(* IEC 61131-3 sources: FACTORY_io/fabrica-viva/etapa-6, 3 files *)

(* ---- fragmento-bloques.st ---- *)
(* ===== Etapa 6 · Bloque de función FB_Muting =====
   La cortina del muelle protege a las personas: si algo la corta, la línea se para. Pero los palés
   tienen que pasar por ella. El muting la anula solo mientras pasa un palé:
   - Empieza si los dos sensores de muting se tapan en orden: primero A y después B (el flanco de
     subida de B con A tapado). Una persona que cruza la cortina no los tapa así.
   - Acaba cuando la carga ha pasado: A y B libres y la cortina despejada.
   - Por seguridad, como mucho 30 s seguidos.
   ZonaSegura := la cortina libre, o el muting activo. *)
FUNCTION_BLOCK FB_Muting
VAR_INPUT
  SensorA : BOOL;       (* sensor de muting antes de la cortina *)
  SensorB : BOOL;       (* sensor de muting, más cerca de la cortina *)
  CortinaLibre : BOOL;  (* salida de seguridad de la cortina: TRUE = nada la corta *)
END_VAR
VAR_OUTPUT
  Activo : BOOL;        (* el muting está anulando la cortina *)
  ZonaSegura : BOOL;    (* se puede trabajar *)
END_VAR
VAR
  (* tus variables internas del bloque *)
END_VAR

(* ---- tu código del bloque ---- *)
END_FUNCTION_BLOCK

(* ---- solucion.st ---- *)
(* Fábrica viva · Etapa 6 · Solución de referencia: enfardado, expedición y cortina de seguridad con muting. *)
FUNCTION_BLOCK FB_Cola
VAR_INPUT
  Meter : BOOL;
  Valor : DINT;
  Sacar : BOOL;
END_VAR
VAR_OUTPUT
  Primero : DINT;
  Cantidad : INT;
END_VAR
VAR
  Datos : ARRAY[0..15] OF DINT;
  i : INT;
END_VAR

(* Sacar desplaza todo un puesto hacia la cabeza; meter escribe detrás del último. *)
IF Sacar AND Cantidad > 0 THEN
  FOR i := 0 TO 14 DO
    Datos[i] := Datos[i + 1];
  END_FOR;
  Cantidad := Cantidad - 1;
END_IF;
IF Meter AND Cantidad < 16 THEN
  Datos[Cantidad] := Valor;
  Cantidad := Cantidad + 1;
END_IF;
IF Cantidad > 0 THEN
  Primero := Datos[0];
ELSE
  Primero := 0;
END_IF;
END_FUNCTION_BLOCK

FUNCTION_BLOCK FB_Muting
VAR_INPUT
  SensorA : BOOL;
  SensorB : BOOL;
  CortinaLibre : BOOL;
END_VAR
VAR_OUTPUT
  Activo : BOOL;
  ZonaSegura : BOOL;
END_VAR
VAR
  SubeB : R_TRIG;
  Limite : TON;
END_VAR

(* El muting empieza solo si los dos sensores se tapan en orden, A y luego B, como hace un palé al
   llegar; una persona que cruza la cortina no los tapa así. Acaba cuando la carga ha pasado: los dos
   sensores libres y la cortina despejada. Con un tiempo máximo, por si se queda algo a medias. *)
SubeB(CLK := SensorB);
IF SubeB.Q AND SensorA THEN
  Activo := TRUE;
END_IF;
IF Activo AND NOT SensorA AND NOT SensorB AND CortinaLibre THEN
  Activo := FALSE;
END_IF;
Limite(IN := Activo, PT := T#30s);
IF Limite.Q THEN
  Activo := FALSE;
END_IF;
ZonaSegura := CortinaLibre OR Activo;
END_FUNCTION_BLOCK

FUNCTION_BLOCK FB_Paletizado
VAR_INPUT
  Habilitar : BOOL;
  CajaLista : BOOL;
  PaleListo : BOOL;
  RobotListo : BOOL;
  Reiniciar : BOOL;
END_VAR
VAR_OUTPUT
  Trabajo : INT;
  Ejecutar : BOOL;
  Paso : INT;
  Colocadas : INT;
  Total : INT;
  PaleLleno : BOOL;
END_VAR

(* Intercambio de señales con el robot: se fija el trabajo, se mantiene Ejecutar hasta que el robot
   avisa de que lo ha empezado (cae RobotListo) y se espera a que vuelva a estar listo. *)
Ejecutar := FALSE;
CASE Paso OF
  0: (* esperando caja y palé *)
    IF Reiniciar THEN
      Colocadas := 0;
    END_IF;
    IF Habilitar AND CajaLista AND PaleListo AND RobotListo AND Colocadas < 8 THEN
      Trabajo := 1;
      Paso := 1;
    END_IF;
  1: (* recoger: orden dada *)
    Ejecutar := TRUE;
    IF NOT RobotListo THEN
      Paso := 2;
    END_IF;
  2: (* recogiendo *)
    IF RobotListo AND Habilitar THEN
      Trabajo := 2 + Colocadas;
      Paso := 3;
    END_IF;
  3: (* dejar en su hueco: orden dada *)
    Ejecutar := TRUE;
    IF NOT RobotListo THEN
      Paso := 4;
    END_IF;
  4: (* dejando y volviendo a reposo *)
    IF RobotListo THEN
      Colocadas := Colocadas + 1;
      Total := Total + 1;
      Paso := 0;
    END_IF;
END_CASE;
PaleLleno := Colocadas >= 8;
END_FUNCTION_BLOCK

FUNCTION_BLOCK FB_Pulmon
VAR_INPUT
  Habilitar : BOOL;
  CajaEnTope : BOOL;
  Permiso : BOOL;
END_VAR
VAR_OUTPUT
  Tope : BOOL;
  Avance : BOOL;
  Salida : BOOL;
  Estado : INT;
  Liberadas : INT;
END_VAR
VAR
  Cerrando : TON;
  Bajando : TON;
END_VAR

CASE Estado OF
  0: (* esperando *)
    IF Habilitar AND CajaEnTope AND Permiso THEN
      Estado := 1;
    END_IF;
  1: (* liberando: rodillos parados (la caja siguiente se queda) y tope abajo hasta que la caja se va *)
    IF NOT CajaEnTope THEN
      Liberadas := Liberadas + 1;
      Estado := 2;
    END_IF;
  2: (* cerrando: tope arriba; los rodillos arrancan cuando ha subido *)
    IF Cerrando.Q THEN
      Estado := 0;
    END_IF;
END_CASE;
(* el temporizador se llama fuera del CASE: así ve siempre su entrada *)
Cerrando(IN := Estado = 2, PT := T#500ms);
Bajando(IN := Estado = 1, PT := T#400ms);
Tope := Estado <> 1;
Avance := Habilitar AND Estado = 0;
(* la cinta de salida espera a que el tope haya bajado del todo antes de llevarse la caja *)
Salida := Habilitar AND NOT (Estado = 1 AND NOT Bajando.Q);
END_FUNCTION_BLOCK

FUNCTION_BLOCK FB_Cinta
VAR_INPUT
  Habilitar : BOOL;
  Presencia : BOOL;
  Rearme : BOOL;
END_VAR
VAR_OUTPUT
  Motor : BOOL;
  Atasco : BOOL;
END_VAR
VAR
  Tapada : TON;
END_VAR

Tapada(IN := Presencia AND Motor, PT := T#3s);
IF Rearme THEN
  Atasco := FALSE;
END_IF;
IF Tapada.Q THEN
  Atasco := TRUE;
END_IF;
Motor := Habilitar AND NOT Atasco;
END_FUNCTION_BLOCK

VAR_INPUT
  Marcha : BOOL;
  Paro : BOOL;
  Seta : BOOL;
  FotocelulaRecepcion : BOOL;
  CajasRecibidas : INT;
END_VAR
VAR_OUTPUT
  CintaRecepcion : BOOL;
  Alimentador : BOOL;
  Baliza : INT;
END_VAR
VAR
  EnMarcha : BOOL;
END_VAR

VAR_INPUT
  Rearme : BOOL;
  FotocelulaAtasco : BOOL;
  LecturaOk : BOOL;
  CodigoCaja : DINT;
  FotocelulaRechazo : BOOL;
  CajasRechazadas : INT;
  CajasFinLinea : INT;
END_VAR
VAR_OUTPUT
  CintaControl : BOOL;
  Desvio : BOOL;
  AlarmaAtasco : BOOL;
END_VAR
VAR
  Control : FB_Cinta;
  Leida : R_TRIG;
  Llega : R_TRIG;
  SinEtiqueta : BOOL;
  Pendiente : BOOL;
  Retardo : TON;
  Empuje : TP;
END_VAR

VAR_INPUT
  FotocelulaExpres : BOOL;
  FotocelulaDevol : BOOL;
  CajasExpres : INT;
  CajasDevueltas : INT;
  CajasPedidos : INT;
END_VAR
VAR_OUTPUT
  CintaClasificacion : BOOL;
  DesvioExpres : BOOL;
  DesvioDevol : BOOL;
END_VAR
VAR
  ColaA : FB_Cola;
  ColaB : FB_Cola;
  CodigoEnA : DINT;
  LlegaA : R_TRIG;
  LlegaB : R_TRIG;
  PendienteA : BOOL;
  PendienteB : BOOL;
  RetardoA : TON;
  RetardoB : TON;
  EmpujeA : TP;
  EmpujeB : TP;
END_VAR

VAR_INPUT
  FotocelulaEntradaPulmon : BOOL;
  FotocelulaLleno : BOOL;
  FotocelulaTope : BOOL;
  FotocelulaSalidaPulmon : BOOL;
  CajasAPaletizar : INT;
END_VAR
VAR_OUTPUT
  RodillosPulmon : BOOL;
  TopePulmon : BOOL;
  CintaSalidaPulmon : BOOL;
  PulmonLleno : BOOL;
END_VAR
VAR
  Pulmon : FB_Pulmon;
  Ritmo : TON;
  LlenoTapada : TON;
  LlenoLibre : TON;
END_VAR

VAR_INPUT
  FotocelulaPicking : BOOL;
  PalePresente : BOOL;
  PaleEnDispensador : BOOL;
  DispensadorOcupado : BOOL;
  RobotListo : BOOL;
  SalidaPales : INT;
END_VAR
VAR_OUTPUT
  RodillosPale : BOOL;
  TopePale : BOOL;
  DarPale : BOOL;
  RobotTrabajo : INT;
  RobotEjecutar : BOOL;
  RobotHabilitado : BOOL;
  CajasPaletizadas : INT;
  PalesCompletos : INT;
END_VAR
VAR
  Paletizado : FB_Paletizado;
  PasoPale : INT;
  CajaQuieta : TON;
  Asentado : TON;
  Fuera : TON;
END_VAR

VAR_INPUT
  PaleEnEnfardadora : BOOL;
  EnfardadoraOcupada : BOOL;
  EnfardadoHecho : BOOL;
  CortinaLibre : BOOL;
  MutingA : BOOL;
  MutingB : BOOL;
  PaleEnMuelle : BOOL;
  SalidaExpedicion : INT;
END_VAR
VAR_OUTPUT
  RodillosEnfardado : BOOL;
  Enfardar : BOOL;
  EnfardadoraHabilitada : BOOL;
  RodillosExpedicion : BOOL;
  LamparaMuting : BOOL;
  AlarmaCortina : BOOL;
  PalesExpedidos : INT;
END_VAR
VAR
  Muting : FB_Muting;
  PasoEnf : INT;
  Salido : TON;
  MuelleOcupado : TOF;
  LlegaMuelle : F_TRIG;
END_VAR

(* Etapas 1 y 2 *)
EnMarcha := (Marcha OR EnMarcha) AND NOT Paro AND Seta AND NOT AlarmaAtasco AND NOT AlarmaCortina;
CintaRecepcion := EnMarcha;
Alimentador := EnMarcha AND NOT PulmonLleno;
Control(Habilitar := EnMarcha, Presencia := FotocelulaAtasco, Rearme := Rearme);
CintaControl := Control.Motor;
AlarmaAtasco := Control.Atasco;
IF NOT Seta OR AlarmaCortina THEN
  Baliza := 4;
ELSIF AlarmaAtasco THEN
  Baliza := 6;
ELSIF EnMarcha AND PulmonLleno THEN
  Baliza := 3;
ELSIF EnMarcha THEN
  Baliza := 1;
ELSE
  Baliza := 2;
END_IF;
Leida(CLK := LecturaOk);
IF Leida.Q THEN
  SinEtiqueta := CodigoCaja = 0;
END_IF;
Llega(CLK := FotocelulaRechazo);
IF Llega.Q AND SinEtiqueta AND EnMarcha THEN
  Pendiente := TRUE;
END_IF;
Retardo(IN := Pendiente, PT := T#450ms);
IF Retardo.Q OR NOT EnMarcha THEN
  Pendiente := FALSE;
END_IF;
Empuje(IN := Retardo.Q, PT := T#600ms);
Desvio := Empuje.Q AND EnMarcha;

(* Etapa 3. Primero se detectan las llegadas; después se decide con la cabeza de cada cola (el código de la
   caja que acaba de llegar) y por último se actualizan las colas, cada una con una sola llamada por ciclo. *)
CintaClasificacion := EnMarcha;
LlegaB(CLK := FotocelulaDevol);
LlegaA(CLK := FotocelulaExpres);
IF LlegaB.Q AND ColaB.Primero = 104 THEN
  PendienteB := TRUE;
END_IF;
CodigoEnA := ColaA.Primero;
IF LlegaA.Q AND CodigoEnA = 103 THEN
  PendienteA := TRUE;
END_IF;
(* la caja que pasa el empujador exprés sin desviarse entra en la cola del tramo siguiente *)
ColaB(Meter := LlegaA.Q AND ColaA.Cantidad > 0 AND CodigoEnA <> 103, Valor := CodigoEnA, Sacar := LlegaB.Q);
ColaA(Meter := Leida.Q AND CodigoCaja <> 0, Valor := CodigoCaja, Sacar := LlegaA.Q);

RetardoA(IN := PendienteA, PT := T#450ms);
IF RetardoA.Q OR NOT EnMarcha THEN
  PendienteA := FALSE;
END_IF;
EmpujeA(IN := RetardoA.Q, PT := T#600ms);
DesvioExpres := EmpujeA.Q AND EnMarcha;
RetardoB(IN := PendienteB, PT := T#450ms);
IF RetardoB.Q OR NOT EnMarcha THEN
  PendienteB := FALSE;
END_IF;
EmpujeB(IN := RetardoB.Q, PT := T#600ms);
DesvioDevol := EmpujeB.Q AND EnMarcha;

(* Etapa 4: el pulmón suelta una caja cada 10 s como mucho, y retiene la descarga si se llena. *)
Ritmo(IN := Pulmon.Estado = 0, PT := T#10s);
(* etapa 5: además, solo con el punto de recogida libre, para no bajar el tope con la cinta de salida parada *)
Pulmon(Habilitar := EnMarcha, CajaEnTope := FotocelulaTope, Permiso := Ritmo.Q AND NOT FotocelulaPicking);
TopePulmon := Pulmon.Tope;
RodillosPulmon := Pulmon.Avance;
LlenoTapada(IN := FotocelulaLleno, PT := T#2s);
LlenoLibre(IN := NOT FotocelulaLleno, PT := T#3s);
IF LlenoTapada.Q THEN
  PulmonLleno := TRUE;
ELSIF LlenoLibre.Q THEN
  PulmonLleno := FALSE;
END_IF;

(* Etapa 5: la cinta de salida lleva cada caja al punto de recogida y espera allí a que el robot la coja. *)
CintaSalidaPulmon := Pulmon.Salida AND NOT FotocelulaPicking;
CajaQuieta(IN := FotocelulaPicking, PT := T#300ms);
RobotHabilitado := EnMarcha;

(* Palés: pedir uno al dispensador, llevarlo al tope, cargarlo y sacarlo lleno. *)
DarPale := FALSE;
RodillosPale := FALSE;
TopePale := TRUE;
CASE PasoPale OF
  0: (* pedir un palé (el dispensador actúa en el flanco de subida) *)
    IF EnMarcha AND NOT DispensadorOcupado THEN
      PasoPale := 1;
    END_IF;
  1:
    DarPale := TRUE;
    IF DispensadorOcupado THEN
      PasoPale := 2;
    END_IF;
  2: (* el dispensador lo deja sobre los rodillos: no se mueven hasta que termina *)
    IF NOT DispensadorOcupado THEN
      PasoPale := 3;
    END_IF;
  3: (* llevarlo hasta el tope *)
    RodillosPale := EnMarcha;
    IF Asentado.Q THEN
      PasoPale := 4;
    END_IF;
  4: (* cargando: lo hace el robot *)
    IF Paletizado.PaleLleno AND Paletizado.Paso = 0 THEN
      PasoPale := 5;
    END_IF;
  5: (* sacar el palé lleno *)
    TopePale := FALSE;
    RodillosPale := EnMarcha;
    IF Fuera.Q THEN
      PalesCompletos := PalesCompletos + 1;
      PasoPale := 0;
    END_IF;
END_CASE;
Asentado(IN := PasoPale = 3 AND PalePresente, PT := T#2s);
Fuera(IN := PasoPale = 5 AND NOT PalePresente, PT := T#3s);

Paletizado(Habilitar := EnMarcha, CajaLista := CajaQuieta.Q, PaleListo := PasoPale = 4, RobotListo := RobotListo,
  Reiniciar := PasoPale <> 4);
RobotTrabajo := Paletizado.Trabajo;
RobotEjecutar := Paletizado.Ejecutar;
CajasPaletizadas := Paletizado.Total;

(* Etapa 6: la cortina del muelle. Si se corta sin muting, alarma: se para la línea y hace falta
   Rearme (con la cortina despejada) y luego Marcha. *)
Muting(SensorA := MutingA, SensorB := MutingB, CortinaLibre := CortinaLibre);
LamparaMuting := Muting.Activo;
IF NOT Muting.ZonaSegura THEN
  AlarmaCortina := TRUE;
ELSIF Rearme THEN
  AlarmaCortina := FALSE;
END_IF;

(* Enfardado: recibir el palé, pararlo bajo el brazo, enfardar y soltarlo. *)
Enfardar := FALSE;
RodillosEnfardado := FALSE;
EnfardadoraHabilitada := EnMarcha;
CASE PasoEnf OF
  0: (* recibir *)
    RodillosEnfardado := EnMarcha;
    IF PaleEnEnfardadora THEN
      PasoEnf := 1;
    END_IF;
  1: (* orden de enfardar (flanco) *)
    Enfardar := TRUE;
    IF EnfardadoraOcupada THEN
      PasoEnf := 2;
    END_IF;
  2: (* enfardando *)
    IF EnfardadoHecho THEN
      PasoEnf := 3;
    END_IF;
  3: (* soltar hacia el muelle *)
    RodillosEnfardado := EnMarcha;
    IF Salido.Q THEN
      PasoEnf := 0;
    END_IF;
END_CASE;
Salido(IN := PasoEnf = 3 AND NOT PaleEnEnfardadora, PT := T#4s);
RodillosExpedicion := EnMarcha;
(* un palé tiene huecos entre sus tacos: la fotocélula parpadea al pasar. Con el TOF, el palé cuenta
   una vez, cuando la fotocélula lleva 1 s libre. *)
MuelleOcupado(IN := PaleEnMuelle, PT := T#1s);
LlegaMuelle(CLK := MuelleOcupado.Q);
IF LlegaMuelle.Q THEN
  PalesExpedidos := PalesExpedidos + 1;
END_IF;

(* ---- fragmento-declaraciones.st ---- *)
(* ===== Etapa 6 · Enfardado y expedición: señales nuevas ===== *)
VAR_INPUT
  PaleEnEnfardadora : BOOL;    (* el palé está centrado bajo el brazo de la enfardadora *)
  EnfardadoraOcupada : BOOL;   (* la enfardadora está trabajando: no muevas sus rodillos *)
  EnfardadoHecho : BOOL;       (* palé enfardado y brazo recogido *)
  CortinaLibre : BOOL;         (* cortina de seguridad del muelle: TRUE = nada la corta *)
  MutingA : BOOL;              (* sensor de muting A *)
  MutingB : BOOL;              (* sensor de muting B *)
  PaleEnMuelle : BOOL;         (* fotocélula del muelle, justo antes del camión *)
  SalidaExpedicion : INT;      (* lo que entra en el camión: cada palé y cada caja cuentan 1 *)
END_VAR
VAR_OUTPUT
  RodillosEnfardado : BOOL;    (* rodillos de la enfardadora *)
  Enfardar : BOOL;             (* orden de enfardar (flanco de subida) *)
  EnfardadoraHabilitada : BOOL;(* la enfardadora solo se mueve con esto a TRUE *)
  RodillosExpedicion : BOOL;   (* rodillos de expedición, hasta el camión *)
  LamparaMuting : BOOL;        (* lámpara de muting de la cortina *)
  AlarmaCortina : BOOL;        (* alguien ha cortado la cortina sin muting *)
  PalesExpedidos : INT;        (* objetivo en directo *)
END_VAR
VAR
  Muting : FB_Muting;          (* tu muting de la cortina *)
  PasoEnf : INT;               (* tu secuencia de enfardado *)
END_VAR
